(*!
<summary>Provides fixed-capacity storage for JSON text.</summary>
<description>
Holds up to 25000 STRING bytes plus the terminator. The alias does not parse or validate JSON.
</description>
*)
(*
SPDX-FileCopyrightText: © 2026 Oleksandr Tiutyk <trofimich@gmail.com>
SPDX-License-Identifier: MIT
License: https://opensource.org/license/mit
*)

TYPE JSON_DOCUMENT : STRING(Parameters.JSON_DOCUMENT_CHAR_SIZE); END_TYPE

(* stored: Version 1.1.0.1
   DUT JSON_DOCUMENT: Id {1c584fbf-bc67-4669-8e1b-884fc72f5a93} *)
